// TIA Portal V21 export
// export: Created 2026-11-10T07:35:23.5631062Z, ExportSetting WithDefaults, DisplayName Totally Integrated Automation Portal, DisplayVersion V21 Update 3, DisplayName STEP 7 Professional, DisplayVersion V21 Update 3, DisplayName STEP 7 Safety, DisplayVersion V21, DisplayName Tech WebApplication, DisplayVersion V21, DisplayName WinCC Basic/Comfort/Advanced, DisplayVersion V21 Update 3, DisplayName WinCC Unified, DisplayVersion V21 Update 3
FUNCTION_BLOCK "FB_Lad_ex156"   // FB58, LAD
{ S7_Optimized_Access := 'TRUE' }
VERSION : 0.1
// stored: AutoNumber true, IsIECCheckEnabled false, IsRetainMemResEnabled false, MemoryReserve 100, SetENOAutomatically false, UDAEnableTagReadback false
   VAR_INPUT
      v_laddr : HW_IO;
      v_ret_val : Int;
   END_VAR
   VAR_OUTPUT
      v_piaddr : UDInt;
      v_picount : UInt;
      v_pqaddr : UDInt;
      v_pqcount : UInt;
   END_VAR
BEGIN

REGION Network 1: RD_ADDR - Determine IO addresses from the hardware identifier
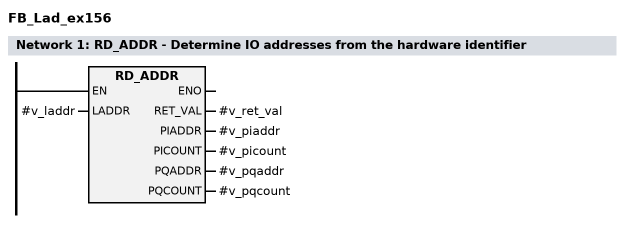
   RUNG wire#powerrail
      RD_ADDR(LADDR := #v_laddr, Ret_Val => #v_ret_val, PIADDR => #v_piaddr, PICount => #v_picount, PQADDR => #v_pqaddr, PQCount => #v_pqcount)
   END_RUNG
   // the same network as SCL:
   #v_ret_val := RD_ADDR(LADDR := #v_laddr,
                         PIADDR => #v_piaddr,
                         PICount => #v_picount,
                         PQADDR => #v_pqaddr,
                         PQCount => #v_pqcount);
END_REGION
END_FUNCTION_BLOCK
